TYPE ST_LightState :
STRUCT
    bValid : BOOL;
    bOn : BOOL;
END_STRUCT
END_TYPE

(* stored: Version 1.1.0.1
   DUT ST_LightState: Id {258a78a9-6fa9-4263-af2a-198b19e334a2} *)
